  # add a "skill" to the robots skillset the control system will send a string with the ls_item and action and here we will look if we have a matching skill to execute
  # the item_modell defines the patterns which have to be used by the robot on multiple racks and or multiple samples in a rackpattern
  # inner pattern is always dependung on the object that has to be moved and the outer pattern is the pattern for the containers where the objects are stored in.
  # if racks have to be handled it is also an inner pattern cause the object to handle is the rack itself
  # create_item(id=0, ls_item="default", frame=p[0,0,0,0,0,0], actionlist=create_action_list([]), item_model=create_item_model(), lm_id=0, description="default")
  # create_item_model(inner=create_pattern(), outer=create_pattern(), description="default")
  # ITEM_MAP.append(create_item(id=1, ls_item="Home", frame=F1_uLM_Home, actionlist=[ActionManipulator.MOVE_TO], description="uLM Move To Home"))
  # ITEM_MAP.append(create_item(id=2, ls_item="InputStation", frame=F2_uLM_Input, actionlist=[ActionManipulator.PICK, ActionManipulator.PLACE], item_model=create_item_model(inner=Patterns.INPUT), description="uLM Pick and Place samples from Input"))
  # ITEM_MAP.append(create_item(id=3, ls_item="InputCapture", frame=F3_Cap_Input, actionlist=[ActionCamera.INSPECT, ActionManipulator.MOVE_TO], description="uLM Inspect samples from Input and Move To Capture Position"))
  # ITEM_MAP.append(create_item(id=4, ls_item="Bin", frame=F4_uLM_Bin, actionlist=[ActionManipulator.PLACE], description="uLM Place Cap to Bin"))
  # ITEM_MAP.append(create_item(id=5, ls_item="StationaryGripper", frame=F5_uLM_Gripper, actionlist=[ActionManipulator.PICK, ActionManipulator.PLACE, ActionManipulator.DECAP, ActionManipulator.MOVE_TO, ActionManipulator.GRASP, ActionManipulator.RELEASE], description=" uLM stationary gripper"))
  # ITEM_MAP.append(create_item(id=6, ls_item="CobasRack", frame=F6_uLM_Cobas_R, actionlist=[ActionManipulator.PICK, ActionManipulator.PLACE], item_model=create_item_model(outer=Patterns.COBAS_MAGAZINE), description="uLM Cobas Racks Pick and Place"))
  # ITEM_MAP.append(create_item(id=7, ls_item="CobasMagazine", frame=F7_uLM_Coba_Mag, actionlist=[ActionManipulator.PICK, ActionManipulator.PLACE], item_model=create_item_model(inner=Patterns.COBAS, outer=Patterns.COBAS_MAGAZINE), description="uLM Cobas Magazine Samples Pick and Place"))
  # ITEM_MAP.append(create_item(id=8, ls_item="DetectCobasRacks", frame=F8_Cap_Cobas_LM, actionlist=[ActionCamera.DETECT_OBJECTS, ActionManipulator.MOVE_TO], lm_id=2, description="uLM Cobas Rack Detection and Move To Capture"))
  # ITEM_MAP.append(create_item(id=9, ls_item="TaraMagazine", frame=F9_uLM_Tara, actionlist=[ActionManipulator.PICK, ActionManipulator.PLACE], item_model=create_item_model(inner=Patterns.TARA), description="uLM Centrifuge Tara Pick and Place"))
  # ITEM_MAP.append(create_item(id=10, ls_item="CentrifugeCapture", frame=F10_Cap_CF, actionlist=[ActionManipulator.MOVE_TO, ActionCamera.DETECT], lm_id=1, description="Centrifuge Device Move to Capture Pos and Detect Landmarks"))
  # ITEM_MAP.append(create_item(id=11, ls_item="Centrifuge", frame=F11_CF_PiPl, actionlist=[ActionManipulator.PICK, ActionManipulator.PLACE], description="Centrifuge Device Rack Pick and Place"))
  # ITEM_MAP.append(create_item(id=12, ls_item="CentrifugeMagazine", frame=F12_uLM_CF_Mag, actionlist=[ActionManipulator.PICK, ActionManipulator.PLACE], item_model=create_item_model(inner=Patterns.CENTRIFUGE, outer=Patterns.CENTRIFUGE_MAGAZINE), description=" uLM Centrifuge Magazin Pick and Place"))
  # ITEM_MAP.append(create_item(id=13, ls_item="CentrifugeRack", frame=F13_uLM_CF_R, actionlist=[ActionManipulator.PICK, ActionManipulator.PLACE], item_model=create_item_model(outer=Patterns.CENTRIFUGE_MAGAZINE), description="uLM Centrifuge Magazin Pick and Place Racks"))
  # ITEM_MAP.append(create_item(id=14, ls_item="DailyArchive", frame=F14_uLM_Archive, actionlist=[ActionManipulator.PICK, ActionManipulator.PLACE], item_model=create_item_model(inner=Patterns.ARCHIVE), description="uLM Pick and Place samples from Archive Rack"))
  # ITEM_MAP.append(create_item(id=15, ls_item="NokRack", frame=F15_uLM_Nok, actionlist=[ActionManipulator.PICK, ActionManipulator.PLACE], item_model=create_item_model(inner=Patterns.NOK), description="uLM Pick and Place samples from Nok Rack"))
  # ITEM_MAP.append(create_item(id=16, ls_item="CobasInput", frame=F16_Cobas_Input, actionlist=[ActionManipulator.PLACE], description="uLM Place Cobasrack in Cobas Device"))
  # ITEM_MAP.append(create_item(id=17, ls_item="CobasInputCapture", frame=F17_Cobas_Cap, actionlist=[ActionCamera.DETECT, ActionManipulator.MOVE_TO], lm_id=3, description="uLM Place Cobasrack in Cobas Device"))
  # ITEM_MAP.append(create_item(id=18, ls_item="XN550Input", frame=F18_XN550_Input, actionlist=[ActionManipulator.PICK, ActionManipulator.PLACE], item_model=create_item_model(inner=Patterns.SYSMEX_XN550, outer=Patterns.DRAWER_XN550), lm_id=4, description="uLM Pick and Place Samples in or out of XN550 Racks"))
  # ITEM_MAP.append(create_item(id=19, ls_item="XN550Capture", frame=F19_XN550_Cap, actionlist=[ActionCamera.DETECT, ActionManipulator.MOVE_TO], lm_id=4, description="uLM Move To and Capture LM XN550"))
  # ITEM_MAP.append(create_item(id=20, ls_item="XN550Drawer", frame=F20_XN550_Draw, actionlist=[ActionManipulator.DRAWER_OPEN, ActionManipulator.DRAWER_CLOSE], item_model=create_item_model(inner=Patterns.DRAWER_XN550), lm_id=4, description="uLM Open and close Drawer XN550"))
  # ITEM_MAP.append(create_item(id=21, ls_item="XN550Button", frame=F21_XN550_Btn, actionlist=[ActionManipulator.PUSH], lm_id=4, description="uLM Push XN550 Button"))
  # ITEM_MAP.append(create_item(id=22, ls_item="AMR", frame=p[0,0,0,0,0,0], actionlist=[ActionAMR.READ, ActionAMR.LOAD_MISSION, ActionAMR.START_MISSION, ActionAMR.NAVIGATE, ActionAMR.ACKNOWLEDGE], description="all AMR actions"))



  # ITEM_MAP.append(create_item(id=31, ls_item="TestLM", frame=TestLM, actionlist=[ActionManipulator.PICK, ActionManipulator.PLACE], item_model=create_item_model(inner=Rack.SYSMEX_CS2500), lm_id=5, description="LM Test"))
  # Fills the Vision Config List with Projectrelated Data
  # workspaceid and skillid are highly robominds related so probably will not stay like this in the future
  # sample detection: dx and dy are used to calculate the positions in a rack and given by the offset which will be applied in order to assign the sample to a place in the rack
  # create_vision_config(workspace_id="", skill_id="", item_id=-1, capture_pos=p[0,0,0,0,0,0], dx=0, dy=0, target_origin=p[0,0,0,0,0,0], selector="default", description="default")
  # VISION_CONFIG_MAP.append(create_vision_config(workspace_id="96017791-f581-4e9e-93da-6951695fccc8", skill_id="8885cfe1-6784-4293-bd26-52ebdc67bf95", capture_pos=F10_Cap_CF, target_origin=p[0,0,0,0,0,0], item_id=11, description="LM Detect CF"))
  # VISION_CONFIG_MAP.append(create_vision_config(workspace_id="96017791-f581-4e9e-93da-6951695fccc8", skill_id="8885cfe1-6784-4293-bd26-52ebdc67bf95", capture_pos=F8_Cap_Cobas_LM, target_origin=p[0,0,0,0,0,0], item_id=8, description="LM Detect Cobas Racks"))
  # VISION_CONFIG_MAP.append(create_vision_config(workspace_id="8f0ad01c-dc36-4fdd-b295-0b6b4a38b89a", skill_id="afdc9e13-ea83-40d6-a805-bb041453d2e5", capture_pos=F3_Cap_Input, target_origin=F2_uLM_Input, item_id=3, description="Lab Solution Input Capture"))
  # VISION_CONFIG_MAP.append(create_vision_config(workspace_id="96017791-f581-4e9e-93da-6951695fccc8", skill_id="8885cfe1-6784-4293-bd26-52ebdc67bf95", capture_pos=F19_XN550_Cap, target_origin=F18_XN550_Input, item_id=18, description="Input XN550"))
  # VISION_CONFIG_MAP.append(create_vision_config(workspace_id="96017791-f581-4e9e-93da-6951695fccc8", skill_id="8885cfe1-6784-4293-bd26-52ebdc67bf95", capture_pos=F19_XN550_Cap, target_origin=POS_Z, item_id=19, description="LM Detect XN550F"))
  # VISION_CONFIG_MAP.append(create_vision_config(workspace_id="96017791-f581-4e9e-93da-6951695fccc8", skill_id="8885cfe1-6784-4293-bd26-52ebdc67bf95", capture_pos=F10_Cap_CF, target_origin=POS_Z, item_id=10, description="LM Detect CF"))
  # VISION_CONFIG_MAP.append(create_vision_config(workspace_id="96017791-f581-4e9e-93da-6951695fccc8", skill_id="8885cfe1-6784-4293-bd26-52ebdc67bf95", capture_pos=F19_XN550_Cap, target_origin=F20_XN550_Draw, item_id=20, description="Drawer XN550"))
  # VISION_CONFIG_MAP.append(create_vision_config(workspace_id="96017791-f581-4e9e-93da-6951695fccc8", skill_id="8885cfe1-6784-4293-bd26-52ebdc67bf95", capture_pos=F19_XN550_Cap, target_origin=F21_XN550_Btn, item_id=21, description="Button XN550"))
  # VISION_CONFIG_MAP.append(create_vision_config(workspace_id="96017791-f581-4e9e-93da-6951695fccc8", skill_id="8885cfe1-6784-4293-bd26-52ebdc67bf95", capture_pos=TestLMCap, target_origin=p[0,0,0,0,0,0], item_id=30, description="Button XN550"))
  # VISION_CONFIG_MAP.append(create_vision_config(workspace_id="96017791-f581-4e9e-93da-6951695fccc8", skill_id="8885cfe1-6784-4293-bd26-52ebdc67bf95", capture_pos=TestLMCap, target_origin=TestLM, item_id=31, description="Button XN550"))

  # VISION_CONFIG_MAP.append(create_vision_config(workspace_id="96017791-f581-4e9e-93da-6951695fccc8", skill_id="8885cfe1-6784-4293-bd26-52ebdc67bf95", target_origin=p[0,0,0,0,0,0], item_id=11, description="LM Detect CF"))
  # VISION_CONFIG_MAP.append(create_vision_config(workspace_id="96017791-f581-4e9e-93da-6951695fccc8", skill_id="8885cfe1-6784-4293-bd26-52ebdc67bf95", target_origin=p[0,0,0,0,0,0], item_id=8, description="LM Detect Cobas Racks"))
  # VISION_CONFIG_MAP.append(create_vision_config(workspace_id="8f0ad01c-dc36-4fdd-b295-0b6b4a38b89a", skill_id="afdc9e13-ea83-40d6-a805-bb041453d2e5", target_origin=F2_uLM_Input, item_id=3, description="Lab Solution Input Capture"))
  # VISION_CONFIG_MAP.append(create_vision_config(workspace_id="96017791-f581-4e9e-93da-6951695fccc8", skill_id="8885cfe1-6784-4293-bd26-52ebdc67bf95", target_origin=F18_XN550_Input, item_id=18, description="Input XN550"))
  # VISION_CONFIG_MAP.append(create_vision_config(workspace_id="96017791-f581-4e9e-93da-6951695fccc8", skill_id="8885cfe1-6784-4293-bd26-52ebdc67bf95", target_origin=POS_Z, item_id=19, description="LM Detect XN550F"))
  # VISION_CONFIG_MAP.append(create_vision_config(workspace_id="96017791-f581-4e9e-93da-6951695fccc8", skill_id="8885cfe1-6784-4293-bd26-52ebdc67bf95", target_origin=POS_Z, item_id=10, description="LM Detect CF"))
  # VISION_CONFIG_MAP.append(create_vision_config(workspace_id="96017791-f581-4e9e-93da-6951695fccc8", skill_id="8885cfe1-6784-4293-bd26-52ebdc67bf95", target_origin=F20_XN550_Draw, item_id=20, description="Drawer XN550"))
  # VISION_CONFIG_MAP.append(create_vision_config(workspace_id="96017791-f581-4e9e-93da-6951695fccc8", skill_id="8885cfe1-6784-4293-bd26-52ebdc67bf95", target_origin=F21_XN550_Btn, item_id=21, description="Button XN550"))
  # VISION_CONFIG_MAP.append(create_vision_config(workspace_id="96017791-f581-4e9e-93da-6951695fccc8", skill_id="8885cfe1-6784-4293-bd26-52ebdc67bf95", target_origin=p[0,0,0,0,0,0], item_id=30, description="Button XN550"))
  # VISION_CONFIG_MAP.append(create_vision_config(workspace_id="96017791-f581-4e9e-93da-6951695fccc8", skill_id="8885cfe1-6784-4293-bd26-52ebdc67bf95", target_origin=TestLM, item_id=31, description="Button XN550"))

  # local inputrack = find_pattern_by_name("INPUT")
  # INSPECT_CONFIG_MAP.append(create_inspect_config(item_id=3, dx=inputrack.pattern_width[0]/(inputrack.pattern_size[0]-1), dy=inputrack.pattern_width[1]/(inputrack.pattern_size[1]-1), rack_size=inputrack.pattern_size , description="Input Capture"))
  # # Fills the Landmark List with Projectrelated Data
  # # create_landmark(lm_id=0, marker_id=-1, marker_size=0.1, marker_type="aruco_7x7", capture_pos=p[0,0,0,0,0,0], init_frame=p[0,0,0,0,0,0], search_offset=[0,0,0], actual_frame=p[0,0,0,0,0,0], description="")
  # LANDMARK_MAP.append(create_landmark(lm_id=1, marker_id=3, marker_size=0.1, marker_type="aruco_7x7", capture_pos = F10_Cap_CF, init_frame=p[-0.617789, -0.065471, 0.07918, 0.020983, -0.012695, 1.512066], search_offset=[0.15, 0.15, 0.1], actual_frame=p[-0.617789, -0.065471, 0.07918, 0.020983, -0.012695, 1.512066], description="LM CF Lid"))
  # LANDMARK_MAP.append(create_landmark(lm_id=2, marker_id=-1, marker_size=0.0085, marker_type="aruco_4x4", capture_pos = F8_Cap_Cobas_LM, init_frame=p[0,0,0,0,0,0], search_offset=[0.15, 0.15, 0.1], actual_frame=POS_Z, description="LM Cobas Rack Detection"))
  # LANDMARK_MAP.append(create_landmark(lm_id=3, marker_id=0, marker_size=0.1, marker_type="aruco_7x7", capture_pos = F17_Cobas_Cap, init_frame=p[-0.667,-0.194,0.100,0,0,0], search_offset=[0.15, 0.15, 0.1], actual_frame=POS_Z, description="LM Cobas Cap"))
  # LANDMARK_MAP.append(create_landmark(lm_id=4, marker_id=4, marker_size=0.1, marker_type="aruco_7x7", capture_pos = F19_XN550_Cap, init_frame=p[0.124,-0.976,0.355,-0.008,0.025,3.131], search_offset=[0.15, 0.15, 0.1], actual_frame=p[0,0,0,0,0,0], description="LM XN550 Cap"))
  # LANDMARK_MAP.append(create_landmark(lm_id=5, marker_id=0, marker_size=0.1, marker_type="aruco_7x7", capture_pos = TestLMCap, init_frame=p[-0.49,-0.144,0.092,0,-0.008,0.001], search_offset=[0.15, 0.15, 0.1], actual_frame=POS_Z, description="LM Test"))
  # # Configuration of all movement related parameters
  # # create_movement(id=0, hh_approach=POS_Z, h_approach=POS_Z, approach=POS_Z, h_target=POS_Z, target=POS_Z, retract=POS_Z, h_retract=POS_Z, hh_retract=POS_Z, h_frame=POS_Z, frame=POS_Z, speed=1, acceleration=1, description="default")
  # MOVEMENT_MAP.append(create_movement(description="TestLMCap", frame=TestLMCap, actionlist=[ActionManipulator.MOVE_TO]))
  # MOVEMENT_MAP.append(create_movement(description="TestLM", frame=TestLM, actionlist=[ActionManipulator.PICK,ActionManipulator.PLACE],
  #         approach=p[0,0,0.1,0,0,0],
  #         retract=p[0,0,0.1,0,0,0]))
  # MOVEMENT_MAP.append(create_movement(description="Home - MOVE_TO", frame=F1_uLM_Home, actionlist=[ActionManipulator.MOVE_TO]))
  # MOVEMENT_MAP.append(create_movement(description="Input - PICK&PLACE", frame=F2_uLM_Input, actionlist=[ActionManipulator.PICK,ActionManipulator.PLACE],
  #         approach=p[0,0,0.1,0,0,0],
  #         retract=p[0,0,0.1,0,0,0]))
  # MOVEMENT_MAP.append(create_movement(description="Capture Input - MOVE_TO", frame=F3_Cap_Input, actionlist=[ActionManipulator.MOVE_TO]))
  # MOVEMENT_MAP.append(create_movement(description="BIN - PLACE", frame=F4_uLM_Bin, actionlist=[ActionManipulator.PLACE],
  #         approach=p[0,0,0.1,0,0,0],
  #         retract=p[0,0,0.1,0,0,0]))
  # MOVEMENT_MAP.append(create_movement(description="Gripper - Move To", frame=F5_uLM_Gripper, actionlist=[ActionManipulator.MOVE_TO],
  #         approach=p[0,0,0.1,0,0,0]))
  # MOVEMENT_MAP.append(create_movement(description="Gripper - Pick", frame=F5_uLM_Gripper, actionlist=[ActionManipulator.PICK],
  #         retract=p[0,0,0.1,0,0,0]))
  # MOVEMENT_MAP.append(create_movement(description="Gripper - Place", frame=F5_uLM_Gripper, actionlist=[ActionManipulator.PLACE],
  #         approach=p[0,0,0.1,0,0,0]))
  # MOVEMENT_MAP.append(create_movement(description="CobasRack Pick & Place", frame=F6_uLM_Cobas_R, actionlist=[ActionManipulator.PICK,ActionManipulator.PLACE],
  #         approach=p[0,0,0.1,0,0,0],
  #         target=p[0,0,0,0,0,d2r(90)],
  #         retract=p[0,0,0.1,0,0,0]))
  # MOVEMENT_MAP.append(create_movement(description="CobasMagazine Pick & Place", frame=F7_uLM_Coba_Mag, actionlist=[ActionManipulator.PICK,ActionManipulator.PLACE],
  #         approach=p[0,0,0.1,0,0,0],
  #         target=p[0,0,0,0,0,-d2r(90)],
  #         retract=p[0,0,0.1,0,0,0]))
  # MOVEMENT_MAP.append(create_movement(description="Capture Position Cobas Landmarks", frame=F8_Cap_Cobas_LM, actionlist=[ActionManipulator.MOVE_TO]))
  # MOVEMENT_MAP.append(create_movement(description="TaraMagazine - PICK & PLACE", frame=F9_uLM_Tara, actionlist=[ActionManipulator.PICK,ActionManipulator.PLACE],
  #         approach=p[0,0,0.13,0,0,0],
  #         target=p[0,0,0,0,0,-d2r(90)],
  #         retract=p[0,0,0.13,0,0,0]))
  # MOVEMENT_MAP.append(create_movement(description="Capture Position - Centrifuge LM", frame=F10_Cap_CF,actionlist=[ActionManipulator.MOVE_TO]))
  # MOVEMENT_MAP.append(create_movement(description="Pick and Place Racks - Centrifuge Lid", frame=F11_CF_PiPl, actionlist=[ActionManipulator.PICK,ActionManipulator.PLACE],
  #         approach=p[0,0,0.3,0,0,0],
  #         retract=p[0,0,0.3,0,0,0]))
  # MOVEMENT_MAP.append(create_movement(description="Pick and Place Samples - Centrifuge on uLM", frame=F12_uLM_CF_Mag, actionlist=[ActionManipulator.PICK,ActionManipulator.PLACE],
  #         approach=p[0,0,0.13,0,0,0],
  #         retract=p[0,0,0.13,0,0,0]
  #         ))
  # MOVEMENT_MAP.append(create_movement(description="Pick and Place Racks - Centrifuge on uLM", frame=F13_uLM_CF_R, actionlist=[ActionManipulator.PICK,ActionManipulator.PLACE],
  #         approach=p[0,0,0.15,0,0,0],
  #         retract=p[0,0,0.15,0,0,0]
  #         ))

  # MOVEMENT_MAP.append(create_movement(description="Pick and Place Samples XN550 Racks in Device", frame=F18_XN550_Input, actionlist=[ActionManipulator.PICK,ActionManipulator.PLACE],
  #         approach=p[0,0,0.1,0,0,0],
  #         target = p[0,0,0,0,0,d2r(90)],
  #         retract=p[0,0,0.1,0,0,0]
  #         ))
  # MOVEMENT_MAP.append(create_movement(description="Capture LM XN550", frame=F19_XN550_Cap, actionlist=[ActionManipulator.MOVE_TO]))
  # MOVEMENT_MAP.append(create_movement(description="Open XN550 Drawer ", frame=F20_XN550_Draw, actionlist=[ActionManipulator.DRAWER_OPEN],
  #         h_approach=p[0.07,0,0.1,0,0,0],
  #         approach=p[0,0,0.1,0,0,0],
  #         target = p[0,0,0,0,0,d2r(90)],
  #         retract=p[0.07,0,0,0,0,0],
  #         h_retract=p[0.07,0,0.1,0,0,0]
  #         ))
  # MOVEMENT_MAP.append(create_movement(description="Close XN550 Drawer ", frame=F20_XN550_Draw, actionlist=[ActionManipulator.DRAWER_CLOSE],
  #         h_approach=p[0.07,0,0.1,0,0,0],
  #         approach=p[0.07,0,0,0,0,0],
  #         target = p[0,0,0,0,0,d2r(90)],
  #         retract=p[0,0,0.1,0,0,0],
  #         h_retract=p[0.07,0,0.1,0,0,0]
  #         ))
  # MOVEMENT_MAP.append(create_movement(description="Push XN550 Button ", frame=F21_XN550_Btn, actionlist=[ActionManipulator.PUSH],
  #         approach=p[0,0,0.15,0,0,0],
  #         retract=p[0,0,0.15,0,0,0]
  #         ))
  # MOVEMENT_MAP.append(create_movement(description="Capture Position 2 Input", frame=F_Cap_Input2,actionlist=[ActionManipulator.MOVE_TO]))



  $ 19 "Script: SCRIPT Objects V0.1.script"
  #*****************************************************
  # customer          :   INTERNAL
  # project name      :
  #****************************************************
  # controller        :   UR
  # software          :   5.17.3
  #****************************************************
  # author            :   P. Koehnke
  # Copyright (c)     :   United Robotics Group
  #                       An der Riede 2
  #                       28816 Stuhr
  #                       Germany
  #****************************************************
  # description       :   object database
  # version:      	:   0.1
  # created           :   09.10.2024
  # updated           :
  #****************************************************
  # modifications     :
  #
  # date              :
  # name              :
  # reason            :
  #****************************************************

  def create_object_2(id=0, name="", type=0, dimension=struct(length=0, width=0, height=0, diameter=0), gripper_offset=p[0,0,0,0,0,0]):
      return struct(id=id, name=name, type=type, dimension=dimension, gripper_offset=gripper_offset)
  end

  OBJ = create_object_2()
  OBJs = make_list(0, create_object_2(), 50)

  OBJs.append(create_object_2(id=1, name="rack centrifuge", type=1, dimension=struct(length=0, width=0, height=0.106, diameter=0.020), gripper_offset=p[0,0,0.095,0,0,2.356]))
  OBJs.append(create_object_2(id=2, name="sample tube 1", type=2, dimension=struct(length=0, width=0, height=0.106, diameter=0.015), gripper_offset=p[0,0,0,0,0,0]))
  OBJs.append(create_object_2(id=3, name="rack sarstedt", type=3, dimension=struct(length=0, width=0, height=0.100, diameter=0.020), gripper_offset=p[0,0,0,0,0,0]))
  OBJs.append(create_object_2(id=4, name="Lab bottle", type=4, dimension=struct(length=0, width=0, height=0.100, diameter=0.030), gripper_offset=p[0,0,0.2,0,0,0]))
  OBJs.append(create_object_2(id=5, name="Vial", type=5, dimension=struct(length=0, width=0, height=0.100, diameter=0.0275), gripper_offset=p[0,0,0,0,0,0]))
  OBJs.append(create_object_2(id=6, name="Container", type=6, dimension=struct(length=0.09, width=0.09, height=0.185, diameter=0.080), gripper_offset=p[0,0,0,0,0,0]))
  OBJs.append(create_object_2(id=7, name="Target_container", type=7, dimension=struct(length=0.06, width=0.06, height=0.134, diameter=0.05), gripper_offset=p[0,0,0,0,0,0]))
  OBJs.append(create_object_2(id=8, name="Spatula", type=8, dimension=struct(length=0.03, width=0.03, height=0.23, diameter=0.05), gripper_offset=p[0,0,0,0,0,0]))
  OBJs.append(create_object_2(id=9, name="rack pipet", type=9, dimension=struct(length=0.03, width=0.03, height=0.23, diameter=0.05), gripper_offset=p[0,0,0,0,0,0]))

  def create_jig_2(id=0, name="", type=0, capacity=0, jig_offset=p[0,0,0,0,0,0]):
      # iformation about used jigs
      return struct(id=id, name=name, type=type, capacity=capacity, jig_offset=jig_offset)
  end

  JIG2 = create_jig_2()
  JIGs = make_list(0, create_jig_2(), 20)

  JIGs.append(create_jig_2(id=1, name="3FG", type=1, capacity=1, jig_offset=p[0,0,0,0,0,0]))
  JIGs.append(create_jig_2(id=2, name="jig input", type=2, capacity=1, jig_offset=p[0,0,0,0,0,-3.927]))
  JIGs.append(create_jig_2(id=3, name="jig output", type=3, capacity=1, jig_offset=p[0,0,0,0,0,0.78]))
  JIGs.append(create_jig_2(id=6, name="jig bin", type=6, capacity=1, jig_offset=p[0,0,0,0,0,0]))
  JIGs.append(create_jig_2(id=7, name="jig sarstedt racks", type=7, capacity=1, jig_offset=p[0,0,-0.02,0,0,0]))
  JIGs.append(create_jig_2(id=8, name="NoK Bin", type=8, capacity=1, jig_offset=p[0,0,0,0,0,0]))
  JIGs.append(create_jig_2(id=9, name="Pick bott jig", type=9, capacity=1, jig_offset=p[0,0,0,0,0,0]))
  JIGs.append(create_jig_2(id=10, name="Place bott jig", type=10, capacity=1, jig_offset=p[0,0,0,0,0,0]))
  JIGs.append(create_jig_2(id=11, name="bottle shake jig", type=11, capacity=1, jig_offset=p[0,0,0,0,0,0]))
  JIGs.append(create_jig_2(id=12, name="Pick Vial jig", type=12, capacity=1, jig_offset=p[0,0,0,0,0,0]))
  JIGs.append(create_jig_2(id=13, name="Place Vial jig", type=13, capacity=1, jig_offset=p[0,0,0,0,0,0]))
  JIGs.append(create_jig_2(id=14, name="Liquid transfer jig", type=14, capacity=1, jig_offset=p[0,0,0,0,0,0]))
  JIGs.append(create_jig_2(id=15, name="Pick station jig", type=15, capacity=1, jig_offset=p[0,0,0,0,0,0]))
  JIGs.append(create_jig_2(id=16, name="Place station jig", type=16, capacity=1, jig_offset=p[0,0,0,0,0,0]))
  JIGs.append(create_jig_2(id=17, name="Weigh station jig", type=17, capacity=1, jig_offset=p[0,0,0,0,0,0]))
  JIGs.append(create_jig_2(id=18, name="Pick station 1", type=18, capacity=1, jig_offset=p[0,0,0,0,0,0]))
  JIGs.append(create_jig_2(id=19, name="Pick station 2", type=19, capacity=1, jig_offset=p[0,0,0,0,0,0]))
  JIGs.append(create_jig_2(id=20, name="Pick station 3", type=20, capacity=1, jig_offset=p[0,0,0,0,0,0]))
  JIGs.append(create_jig_2(id=21, name="Tilt station jig", type=21, capacity=1, jig_offset=p[0,0,0,0,0,0]))
  $ 20 "Script: Tilting.script"
  global g_has_ref = False
  global g_pivot_pose = p[0, 0, 0, 0, 0, 0]
  global g_rel0 = p[0, 0, 0, 0, 0, 0]
  global g_current_angle = 0.0

  hinge_offset = p[0, 0, -0.20, 0, 0, 0]
  global g_rq_ready = False
  global RQ_FORCE = 30
  global RQ_SPEED = 100
  global RQ_GRIP_TIMEOUT = 2.0

  def tilt_init_reference():
  	p_center = get_actual_tcp_pose()
  	g_pivot_pose = pose_trans(p_center, hinge_offset)
  	g_rel0 = pose_trans(pose_inv(g_pivot_pose), p_center)
  	g_current_angle = 0.0
  	g_has_ref = True
  end

  def rq_ensure_ready():
  	if (not g_rq_ready):
  		rq_activate_and_wait()
  		rq_set_force(RQ_FORCE)
  		rq_set_speed(RQ_SPEED)
  		g_rq_ready = True
  	end
  end



  #def rq_open_and_wait():
  	#rq_open()
  	#sleep(0.25)
  #end

  def tilt_to(target_deg):
  	if ( not g_has_ref):
  		tilt_init_reference()
  	end

  	rq_ensure_ready()
  	rq_close_and_wait()

  	angle_mid = (g_current_angle + target_deg)/2.0
  	rad_mid = (angle_mid)*3.1416/180
  	rad_end = target_deg*3.1416/180

  	tilt_mid = p[0,0,0, -rad_mid, 0, 0]
  	tilt_end = p[0,0,0, -rad_end, 0, 0]

  	pose_rel_mid = pose_trans(tilt_mid, g_rel0)
  	pose_rel_end = pose_trans(tilt_end, g_rel0)

  	via_pose = pose_trans(g_pivot_pose, pose_rel_mid)
  	end_pose = pose_trans(g_pivot_pose, pose_rel_end)

  	movec(via_pose, end_pose, a=0.05, v=0.01, r=0.001)

  	rq_open_and_wait()

  	g_current_angle = target_deg
  end


  def tilt_by(delta_deg):
  	tilt_to(g_current_angle + delta_deg)
  end

  def tilt_reset():
  	g_has_ref = False
  end

  $ 21 "Script: recipe_updated.script"
  # ============================================
  # Recipe Dosing URScript (3 powders, sorted A/B/C)
  # - keeps final mixture ratio after 1st overshoot
  # - syncs with Python dashboard via TCP
  # ============================================

  # --------- HANDOFF GLOBALS (used by other skills) ---------
  global Pow_name = ""
  global target_weight = 0.0
  global last_dose_error = 0.0

  # --------- RECIPE STATE ---------
  global powder_names = ["", "", ""]
  global powder_ratios = [0.0, 0.0, 0.0]      # fractions 0..1
  global powder_targets = [0.0, 0.0, 0.0]     # target weights for each powder
  global powder_actuals = [0.0, 0.0, 0.0]     # measured after dosing
  global powder_order  = [0, 1, 2]            # indices, sorted by ascending ratio

  global total_weight = 0.0                   # initial / adjusted total
  global current_powder_index = 0             # index into powder_order
  global ratio_adjusted = False               # did we already adjust after powder 1
  global dose_start_weight = 0.0              # weight at dosing start for each powder

  # --------- FINAL RESULTS (for dashboard) ---------
  # WA/WB/WC = final weights of powders A/B/C after dosing (sorted by ratio)
  global WA = 0.0
  global WB = 0.0
  global WC = 0.0

  # finalPercA/B/C = final percentages of WA/WB/WC wrt adjusted total
  global finalPercA = 0.0
  global finalPercB = 0.0
  global finalPercC = 0.0

  # counter to know which powder we just finished (1 → A, 2 → B, 3 → C)
  global dose_counter = 0


  # =====================================================
  # SORTING HELPERS (BY ASCENDING RATIO)
  # =====================================================

  def swap_order(i, j):
    local temp = powder_order[i]
    powder_order[i] = powder_order[j]
    powder_order[j] = temp
  end

  def sort_powders_by_ratio():
    # bubble-sort style, only 3 elements
    global powder_order = [0, 1, 2]

    if (powder_ratios[powder_order[1]] < powder_ratios[powder_order[0]]):
      swap_order(0, 1)
    end

    if (powder_ratios[powder_order[2]] < powder_ratios[powder_order[1]]):
      swap_order(1, 2)
    end

    if (powder_ratios[powder_order[1]] < powder_ratios[powder_order[0]]):
      swap_order(0, 1)
    end
  end


  # =====================================================
  # TCP SENDING HELPERS (Python dashboard @ 192.168.12.103:3002)
  # =====================================================

  # Send powder labels in sorted A/B/C order
  # A = least %, B = middle %, C = highest %
  def send_powder_labels():
    local A = powder_names[powder_order[0]]
    local B = powder_names[powder_order[1]]
    local C = powder_names[powder_order[2]]

    socket_open("192.168.12.103", 3002)
    local cmd = "SET_LABELS:" + A + ";" + B + ";" + C
    textmsg("Sending labels: ", cmd)
    socket_send_string(cmd)
    sleep(0.2)
    socket_close()
  end

  # Send initial recipe (TOTAL;PA;PB;PC) in sorted order
  # powder_ratios are fractions (0..1), we convert to %
  def send_init_recipe(total_w):
    local rA = powder_ratios[powder_order[0]] * 100
    local rB = powder_ratios[powder_order[1]] * 100
    local rC = powder_ratios[powder_order[2]] * 100

    socket_open("192.168.12.103", 3002)
    local cmd = "SET_INIT:" +
                to_str(total_w) + ";" +
                to_str(rA) + ";" +
                to_str(rB) + ";" +
                to_str(rC)
    textmsg("Sending INIT: ", cmd)
    socket_send_string(cmd)
    sleep(0.2)
    socket_close()
  end

  # Send final recipe:
  # SET_FINAL:ADJ_TOTAL;PA;PB;PC;WA;WB;WC
  # where PA/B/C = finalPercA/B/C, WA/B/C = final weights, adj_total = total_weight
  def send_final_recipe(adj_total):
    socket_open("192.168.12.103", 3002)

    local cmd = "SET_FINAL:" +
                to_str(adj_total) + ";" +
                to_str(finalPercA) + ";" +
                to_str(finalPercB) + ";" +
                to_str(finalPercC) + ";" +
                to_str(WA) + ";" +
                to_str(WB) + ";" +
                to_str(WC)
    textmsg("Sending FINAL: ", cmd)
    socket_send_string(cmd)
    sleep(0.2)
    socket_close()
  end


  # =====================================================
  # FINAL WEIGHT & PERCENTAGE LOGIC
  # =====================================================

  # Call this ONCE after each powder dosing is finished
  # final_weight = w_dosed_total of the just-finished powder
  def record_final_weight_for_current_powder(final_weight):
    dose_counter = dose_counter + 1

    if dose_counter == 1:
      WA = final_weight
      textmsg("Assigned WA (Powder A): ", WA)
    elif dose_counter == 2:
      WB = final_weight
      textmsg("Assigned WB (Powder B): ", WB)
    elif dose_counter == 3:
      WC = final_weight
      textmsg("Assigned WC (Powder C): ", WC)
    else:
      textmsg("WARNING: dose_counter > 3, ignoring extra weight")
    end
  end

  # Compute final percentages from WA/WB/WC and adjusted total
  def compute_final_percentages(adj_total):
    if adj_total <= 0:
      textmsg("ERROR: adj_total <= 0, cannot compute final %")
    else:
      finalPercA = WA / adj_total * 100
      finalPercB = WB / adj_total * 100
      finalPercC = WC / adj_total * 100
      textmsg("Final % A/B/C: ", finalPercA, finalPercB, finalPercC)
    end
  end


  # =====================================================
  # RECIPE INITIALIZATION
  # =====================================================

  # powA/B/C  : strings (e.g. "MCC", "CCS", "MAGNESIUM_STEARATE")
  # total     : initial total weight (g)
  # ratioA/B/C: fractions (0..1), e.g. 0.3, 0.2, 0.5
  def recipe_init(powA, powB, powC, total, ratioA, ratioB, ratioC):
    global powder_names  = [powA, powB, powC]
    global powder_ratios = [ratioA, ratioB, ratioC]
    global total_weight  = total

    global powder_targets = [total*ratioA, total*ratioB, total*ratioC]
    global powder_actuals = [0.0, 0.0, 0.0]

    global current_powder_index = 0
    global ratio_adjusted = False
    global dose_start_weight = 0.0

    dose_counter = 0
    WA = 0.0
    WB = 0.0
    WC = 0.0

    sort_powders_by_ratio()

    # NOTE: you call these from your main flow when you want:
    send_powder_labels()
    send_init_recipe(total)
  end


  # =====================================================
  # POSITION + CAMERA HELPERS (YOUR EXISTING LOGIC)
  # =====================================================

  def get_position_for_powder(Pow_name):
    if pos1_powder == Pow_name:
      return "Position1"
    elif pos2_powder == Pow_name:
      return "Position2"
    elif pos3_powder == Pow_name:
      return "Position3"
    else:
      return -1
    end
  end

  def extract_powder_name(raw_str):
    local idx_open  = str_find(raw_str, "(")
    local idx_close = str_find(raw_str, ")")

    if (idx_open < 0) or (idx_close < 0):
      return raw_str
    end

    local inside = ""
    local i = idx_open + 1
    while i < idx_close:
      inside = str_cat(inside, str_at(raw_str, i))
      i = i + 1
    end

    local idx_comma = str_find(inside, ",")
    if idx_comma < 0:
      return inside
    end

    local powder = ""
    local j = idx_comma + 1
    while j < str_len(inside):
      powder = str_cat(powder, str_at(inside, j))
      j = j + 1
    end

    return powder
  end

  def get_response_from_camera(target):
    movel(target, a=0.1, v=0.12, r=0)
    visor_trigger("1", "3.0", "arm")
    global response = visor_getResponse(1)
  end


  # =====================================================
  # RECIPE STEP SELECTION
  # =====================================================

  # Call recipe_next() before each dosing run.
  # Returns True if a powder exists, False if done.
  def recipe_next():
    if (current_powder_index >= 3):
      return False
    end

    local i = powder_order[current_powder_index]
    global Pow_name = powder_names[i]
    global target_weight = powder_targets[i]

    global powder_position = get_position_for_powder(Pow_name)

    if (Pow_name == "CCS"):
      W_now = 200.0
    elif (Pow_name == "MCC"):
      W_now = 131.0
    else:
      W_now = 100.0
    end

    return True
  end


  # =====================================================
  # DOSING START / END
  # =====================================================

  # Call at the beginning of each powder dosing run
  def dosing_start():
    global dose_start_weight = get_weight()
    global switch_spat_M = True
    global switch_spat_S = True
    global switch_spat_F_S = True
  end

  # Call after dosing is finished for current powder
  def dosing_end():
    local idx = powder_order[current_powder_index]
    local weight_after = get_weight()
    local actual_weight = weight_after - dose_start_weight

    # store actual weight
    local tmp = powder_actuals
    tmp[idx] = actual_weight
    global powder_actuals = tmp

    # save error
    global last_dose_error = actual_weight - powder_targets[idx]

    # store WA/WB/WC in dosing (sorted) order
    record_final_weight_for_current_powder(actual_weight)

    # one-time correction after first powder (ratio preserving)
    if ((current_powder_index == 0) and (not ratio_adjusted)):
      local j = powder_order[1]
      local k = powder_order[2]

      local ratio_first = powder_ratios[idx]
      if (ratio_first > 0.0):
        # new_total = actual / ratio_first
        local new_total = actual_weight / ratio_first
        if (new_total < 0.0):
          new_total = 0.0
        end

        local ttmp = powder_targets
        ttmp[idx] = actual_weight
        ttmp[j]   = new_total * powder_ratios[j]
        ttmp[k]   = new_total * powder_ratios[k]
        global powder_targets = ttmp

        global adj_total = new_total
      end

      global ratio_adjusted = True
    end

    global current_powder_index = current_powder_index + 1
  end

  $ 22 "Script: scooping.script"
  def scooping_init():
  	#global W_FULL = 300.010
  	global H_INNER = 0.15
  	global TCP_to_tip = 0.020
  	global depth_saftey = 0.005
  	global container_height = 0.120
  	global reach_margin = 0.03

  	global angle_min = 18.0
  	global angle_max = 68.0
  	global gain_per_percent = 0.5

  	global level_bias_below_center = 0.020

  	global level = 0.0
  	global tilt_angle_sent = 0.0
  	global w_dosed_total = 0.0
  	global last_scale = 0.0
  	global g_z0_hi = 0.01
  	global g_z100_hi = 0.10
  	global g_z_min = 0.018
  	global g_z_max = 0.150

  	#global g_exp = 0.80
  	#global g_k = 0.03
  	#global g_alpha = 0.7
  	global g_corr_max = 0.010

  	global g_prev_cum_w = -1.0
  	global g_depth_corr = 0.0
  	global spatula_len = 0.17
  	global target_g = 0.0
  	global scoop_ct = 0
  	global error_sum = 0.0
  	global error_sq_sum = 0.0
  	global scoop_g = 0.0
  	global w_dosed_total = 0.0

  	if (Pow_name=="NaCl"):
  		global W_FULL = 625.00
  		global g_exp = 0.80
  		global g_k = 0.03
  		global g_alpha = 0.7
  	elif (Pow_name == "Mannitol"):
  		global W_FULL = 300.00
  		global g_exp = 0.82
  		global g_k = 0.025
  		global g_alpha = 0.6
  	elif (Pow_name == "MCC"):
  		global W_FULL = 280.0
  		global g_exp = 0.82
  		global g_k = 0.035
  		global g_alpha = 0.7
  	elif (Pow_name == "CCS"):
  		global W_FULL = 250.0
  		global g_exp = 0.82
  		global g_k = 0.035
  		global g_alpha = 0.7
  	elif (Pow_name == "Magnesium_stearate"):
  		global W_FULL = 200.0
  		global g_exp = 0.84
  		global g_k = 0.025
  		global g_alpha = 0.6
  	elif (Pow_name == "lactose_fine"):
  		global W_FULL = 330.0
  		global g_exp = 0.84
  		global g_k = 0.025
  		global g_alpha = 0.55
  	else:
  		popup("Unkwon powder type. Using default NaCl settings.", title="Calibration Warning")
  		global W_FULL = 300.0
  		global g_k = 0.03
  		global g_alpha = 0.7
  	end


  end

  def clamp(x, lo, hi):
  	if(x<lo):
  		return lo
  	elif (x>hi):
  		return hi
  	else:
  		return x
  	end
  end

  def compute_level_percent(W_now, weight_value):
  	local delta = weight_value - last_scale
  	if (delta<0.0):
  		delta = 0.0
  	end
  	global w_dosed_total = w_dosed_total + delta
  	last_scale = weight_value

  	local W_eff = W_now-w_dosed_total
  	if (W_eff<W_EMPTY):
  		W_eff = W_EMPTY
  	end

  	level = 100.0* (W_eff -W_EMPTY)/ (W_FULL-W_EMPTY)
  	level = clamp(level,0.0,100.0)

  	return level
  end

  def compute_tilt_deg(level_percent):
  	angle = angle_min + gain_per_percent*(100.0-level_percent)
  	return clamp(angle, angle_min, angle_max)
  end


  def tilt(level_percentage):
  	new_angle = compute_tilt_deg(level_percentage)
  	global angle_rel = new_angle - tilt_angle_sent

  	if my_abs(angle_rel)>2.0:
  		tilt_send(new_angle)
  		global angle_deg = new_angle
  		global tilt_angle_sent = new_angle
  		global p_center = updated_center_pose(p_center_vertical, angle_deg)
  	end

  	if (level<85.0):
  		tilt_send(angle_deg)
  	end
  end

  def compute_scoop_depth(level, cum_w, target_g):
  	if (level >=10.0):
  		ratio = level/100.0
  		corrected = pow(ratio, g_exp)
  		base_z = g_z0_hi + (g_z100_hi - g_z0_hi)*corrected

  	elif (level<10.00 and level>=1.00):
  		z0 = 0.023
  		z100 = 0.140
  		ratio2 = level/100.0
  		base_z = z0 +(z100-z0)*ratio2
  	else:
  		base_z = 0.016
  	end

  	if (g_prev_cum_w<0):
  		g_prev_cum_w = cum_w

  	else:
  		global scoop_g = cum_w-g_prev_cum_w
  		g_prev_cum_w = cum_w

  		e = target_g -scoop_g

  		corr_proposed = g_k*e
  		g_depth_corr = (1.0 -g_alpha)*g_depth_corr + g_alpha*corr_proposed
  		g_depth_corr = clamp(g_depth_corr, -g_corr_max, g_corr_max)
  	end

  	z_tip = base_z - g_depth_corr
  	z_tip = clamp(z_tip, g_z_min, g_z_max)


  	return z_tip
  end

  def my_abs(val):
  	if (val<0):
  		return -val
  	else:
  		return val
  	end
  end


  def select_spatula(Pow_name, level, diff):
  	if (Pow_name == "lactose_fine" or Pow_name== "Magnesium_stearate"):
  		if (level >10.0 and diff>0.6):
  			return "spatula_flat_M"
  		else:
  			return "spatula_flat_S"
  		end

  	elif (Pow_name == "NaCl" and level >10.0 and diff>6.5):
  		return "spatula_L"
  	elif(Pow_name == "NaCl" and level> 10.0 and diff<=6.5):
  		return "spatula_M"
  	elif (Pow_name == "MCC" and level >10.0 and diff>2.0):
  		return "spatula_L"
  	elif(Pow_name == "MCC" and level> 10.0 and diff<=2.0):
  		return "spatula_M"
  	elif ((Pow_name == "Mannitol" or Pow_name == "CCS") and level >10.0 and diff>3.2):
  		return "spatula_L"
  	elif ((Pow_name == "Mannitol" or Pow_name == "CCS") and level >10.0 and diff<=3.2):
  		return "spatula_M"
  	elif( level>1.0 and level <= 10.0):
  		return "spatula_M"
  	else:
  		return "spatula_S"
  	end
  end

  global target_g_table = [
  	"NaCl", "spatula_L", "6.8",
  	"NaCl", "spatula_M", "1.75",
  	"NaCl", "spatula_S", "0.135",

  	"Mannitol", "spatula_L", "3.1",
  	"Mannitol", "spatula_M", "0.9",
  	"Mannitol", "spatula_S", "0.075",

  	"CCS", "spatula_L", "2.5",
  	"CCS", "spatula_M", "0.9",
  	"CCS", "spatula_S", "0.075",

  	"MCC", "spatula_L", "1.8",
  	"MCC", "spatula_M", "0.5",
  	"MCC", "spatula_S", "0.05",

  	"Magnesium_stearate", "spatula_flat_M", "0.5",
  	"Magnesium_stearate", "spatula_flat_S", "0.25",

  	"lactose_fine", "spatula_flat_M", "1.0",
  	"lactose_fine", "spatula_flat_S", "0.7"]

  def get_target_g(Pow_name, spat_name):
  	local i = 0
  	local n = length(target_g_table)
  	while (i < n):
  		if (target_g_table[i] == Pow_name and target_g_table[i+1] == spat_name):
  			return to_num(target_g_table[i+2])
  		end
  		i = i+3
  	end
  	popup("No target_g match for: ", Pow_name, ", ", spatula)

  end
  def auto_tilt_and_scoop(W_now, target_weight, weight_value):
  	level = compute_level_percent(W_now, weight_value)

  	global spatula = select_spatula(Pow_name, level, diff)
  	global target_g = get_target_g(Pow_name, spatula)

  	global scoop_depth = compute_scoop_depth(level, weight_value, target_g)

  	tilt(level)
  	#p_center = get_actual_tcp_pose()

  	if (scoop_ct < 5 and g_prev_cum_w>0.0):
  		#local scoop_g = scoop_g
  		local error = target_g - scoop_g
  		error_sum = error_sum + error
  		error_sq_sum = error_sq_sum + error*error
  		scoop_ct = scoop_ct+1

  		if (scoop_ct==5):
  			local avg_error = error_sum/5.0
  			#local std_dev = sqrt(error_sq_sum/5.0) - (avg_error*avg_error))

  			if (my_abs(avg_error)>1.0):
  				g_k = 0.055
  				g_alpha = 0.85
  			elif (my_abs(avg_error)>0.6):
  				g_k= 0.045
  				g_alpha =0.75
  			elif (my_abs(avg_error)> 0.3):
  				g_k = 0.035
  				g_alpha = 0.65
  			elif (my_abs(avg_error)>0.1):
  				g_k = 0.025
  				g_alpha = 0.55
  			else:
  				g_k = 0.015
  				g_alpha = 0.45
  			end
  		end
  	end

  	scoop_powder(p_center)
  end


  def after_scoop():
  	tilt_send(angle_deg)
  	sleep(0.5)
  	movel(lifted_pose, a=0.05, v=0.2)
  	movel(tilted_pose_in_base, a=0.05, v=0.2)
  	set_analog_out(0,0.4)
  	movel(pose_trans(tilted_pose_in_base, p[-0.01,0,0,0,0,2.0]), a=0.05, v=0.2)
  	set_analog_out(0,0.0)
  	movel(lifted_pose, a=0.05, v=0.2)
  	tilt_to_home()
  end
  $ 23 "Script: dosing.script"
  def vibration_2():
  	set_analog_out(0,0.4)
  	sleep(0.8)
  	set_analog_out(0,0.0)
  	sleep(0.2)
  end

  def vibration_3():
  	set_analog_out(0,0.4)
  	sleep(0.5)
  	set_analog_out(0,0.0)
  	sleep(0.3)
  end

  def vibration_4():
  	set_analog_out(0,0.4)
  	sleep(0.6)
  	set_analog_out(0, 0.0)
  	sleep(0.5)
  end

  def vibration_1():
  	set_analog_out(0,0.4)
  	sleep(1)
  	set_analog_out(0,0.0)
  	sleep(0)
  end

  def move_tilt_in_steps(Pow_center, final_pose, steps):
  	i = 0
  	while i <= steps:
  		ratio = i / steps
  		pose_step = p[Pow_center[0] + ratio * (final_pose[0] - Pow_center[0]), Pow_center[1] + ratio * (final_pose[1] -Pow_center[1]),Pow_center[2] + ratio * (final_pose[2] - Pow_center[2]), Pow_center[3] + ratio * (final_pose[3] - Pow_center[3]), Pow_center[4] + ratio * (final_pose[4] - Pow_center[4]), Pow_center[5] + ratio * (final_pose[5] - Pow_center[5])]
  		movej(pose_step, a=1.2, v=0.15)
  		sleep(0.1)
  		i = i+1
  	end
  end

  def tilt_container(angle):
  	p_center = get_actual_tcp_pose()
  	hinge_offset = p[0,0,-0.23,0,0,0]
  	pivot_pose = pose_trans(p_center, hinge_offset)
  	pose_rel = pose_trans(pose_inv(pivot_pose), p_center)
  	angle_mid = (angle/2.0)*3.1416/180
  	angle_end = angle*3.1416/180
  	tilt_mid = p[0,0,0, -angle_mid, 0, 0]
  	tilt_end = p[0,0,0, -angle_end, 0, 0]
  	pose_rel_mid = pose_trans(tilt_mid, pose_rel)
  	pose_rel_end = pose_trans(tilt_end, pose_rel)
  	via_pose = pose_trans(pivot_pose, pose_rel_mid)
  	end_pose = pose_trans(pivot_pose, pose_rel_end)
  	movec(via_pose, end_pose, a=0.05, v=0.01, r=0.001)
  	p_center = get_actual_tcp_pose()
  end

  def deg2rad(d):
  	return d*3.141592/180
  end

  def map_tilt_to_ry_deg(container_deg):
  	#ry_deg = -0.875*container_deg +87.0
  	#return clamp(ry_deg, 5.0, 80.0)
  	if (Pow_name == "NaCl" or Pow_name == "Mannitol" or Pow_name == "CCS" or Pow_name == "MCC"):
  		if ( level>=10.0):
  			ry_min = 10.0
  			ry_max = 75.0
  		elif (level<10.00 and level >1.00):
  			ry_min = 16.0
  			ry_max = 65.0
  		else:
  			ry_min=17.0
  			ry_max=75.0
  		end
  	else:
  		if ( level>=10.0):
  			ry_min = 0.0
  			ry_max = 65.0
  		elif (level<10.00 and level >1.00):
  			ry_min = 10.0
  			ry_max = 45.0
  		else:
  			ry_min=0.0
  			ry_max=50.0
  		end

  	end
  	local span_count = angle_max -angle_min
  	local span_ry = ry_max - ry_min

  	local t = (container_deg -angle_min)/span_count
  	local ry_deg = ry_max - t*span_ry

  	return clamp(ry_deg, ry_min, ry_max)

  end

  def caluclate_corrections(level):
  	z_high = 0.01
  	z_low = -0.08
  	y_high = -0.01
  	y_low = -0.015

  	scale = (level - 10.0) / (100.0-10.0)

  	global correction_z = z_low + scale*(z_high - z_low)
  	global correction_y = y_low + scale*(y_high -y_low)

  end

  def scoop_powder(p_center):
  	#lift_offset = p[0, 0, 0.05, 0, 0, 0]
  	vibration_voltage = 0.4
  	vibration_time = 3.0
  	diameter = 0.07
  	global scoop_radius_default = 0.0
  	#p_center = center_pose_t


  	if (level >=70.00):
  		approach_offset = p[0.008,0,0.22,0,0,0]
  		lift_offset = p[0, 0, 0.05, 0, 0, 0]
  		caluclate_corrections(level)
  	elif (level >=10.00 and level <70):
  		approach_offset = p[0.008,0,0.22,0,0,0]
  		lift_offset = p[0, 0, 0.15, 0, 0, 0]
  		caluclate_corrections(level)
  	elif (level<10.00 and level >= 1.00):
  		approach_offset = p[0.01,0,0.22,0,0,0]
  		correction_z = -0.08
  		correction_y = -0.01
  		lift_offset = p[0, 0, 0.14, 0, 0, 0]
  	else:
  		approach_offset = p[0.008,0,0.22,0,0,0]
  		correction_z = -0.08
  		correction_y = -0.01
  		lift_offset = p[0, 0, 0.14, 0, 0, 0]
   	end

  	if (spatula == "spatula_L"):
  		global spatula_depth = 0.015
  	elif (spatula == "spatula_M"):
  		global spatula_depth = 0.01
  	elif (spatula == "spatula_S"):
  		global spatula_depth = 0.008
  	elif (spatula == "spatula_flat_M"):
  		global spatula_depth = 0.001
  	elif (spatula == "spatula_flat_S"):
  		global spatula_depth = 0.005
  	end

  	scoop_radius_default = diameter/2 - spatula_depth
  	scoop_entry_pose = pose_trans(p_center, approach_offset)
  	movel(scoop_entry_pose, a=0.1, v=0.25)

  	scoop_start_rel = p[scoop_radius_default, 0, scoop_depth, 0, 0, 0]

  	rot_mid = p[0, 0, 0, 0, 0, 0.785]
  	rot_end = p[0, 0, 0, 0, 0, 1.5708]

  	scoop_via_rel = pose_trans(rot_mid, scoop_start_rel)
  	scoop_end_rel = pose_trans(rot_end, scoop_start_rel)

  	scoop_start_pose = pose_trans(p_center, scoop_start_rel)
  	scoop_via_pose = pose_trans(p_center, scoop_via_rel)
  	scoop_end_pose = pose_trans(p_center, scoop_end_rel)

  	movel(scoop_start_pose, a=0.5, v=0.3)
  	#movel(p_center, a=0.5, v=1.0)
  	#sleep(5.0)

  	if (level<90.0):
  		Rotate()
  	end

  	#movec(scoop_via_pose, scoop_end_pose, a=0.03, v=0.05)
  	movec(scoop_via_pose, scoop_end_pose, a=0.03, v=0.02)
  	#movel(pose_trans(get_actual_tcp_pose(), p[0,0,0,0,0,deg2rad(90.0)]), a=0.03, v=0.05)
  	sleep(1.0)
  	local ry_deg = map_tilt_to_ry_deg(angle_deg)
  	local ry = deg2rad(ry_deg)
  	local end_rel = pose_trans(pose_inv(p_center), scoop_end_pose)
  	local end_rel_tilted = pose_trans(end_rel, p[0, 0, 0, 0, ry, 0])
  	global tilted_pose_in_base = pose_trans(p_center, p[0,correction_y,correction_z,end_rel_tilted[3],end_rel_tilted[4], end_rel_tilted[5]])
  	global tilted_pose_in_base = pose_trans(tilted_pose_in_base, p[0, 0, spatula_len, 0, 0, 0])

  	if (Pow_name == "lactose_fine" or Pow_name == "Magnesium_sterate"):
  		tilt_send((angle_deg+5))
  	end
  	movel(tilted_pose_in_base, a=0.03, v=0.1)

  	if (Pow_name == "lactose_fine" or Pow_name == "Magnesium_sterate"):
  		tilt_send((angle_deg-5))
  	end

  	if (spatula=="spatula_flat_S" or spatula=="spatula_S"):
  		vibration_3()
  	else:
  		set_analog_out(0, vibration_voltage)
  	end
  	if (Pow_name=="Mannitol" or Pow_name =="NaCl"):
  		local n=1.4
  	else:
  		local n=1.5
  	end
  	local ry_level = deg2rad(ry_deg/n)
  	local end_rel_tilted_level = pose_trans(end_rel, p[0, 0, 0, 0, ry_level, 0])
  	local level_tilted_pose_in_base = pose_trans(p_center, p[0,correction_y,correction_z,end_rel_tilted_level[3],end_rel_tilted_level[4], end_rel_tilted_level[5]])
  	local level_tilted_pose_in_base = pose_trans(level_tilted_pose_in_base, p[0, 0, spatula_len, 0, 0, 0])

  	movel(level_tilted_pose_in_base, a=0.03, v=0.1)
  	#if (level>70.0):
  		#sleep(1.0)
  	#end
  	sleep(1.0)
  	#sleep(vibration_time)

  	movel(tilted_pose_in_base, a=0.03, v=0.1)
  	set_analog_out(0, 0.0)

  	tilt_pose_rel = pose_trans(pose_inv(p_center), tilted_pose_in_base)

  	lifted_pose_rel = pose_trans(lift_offset, tilt_pose_rel)

  	global lifted_pose = pose_trans(p_center, lifted_pose_rel)
  	movel(lifted_pose, a=0.03, v=0.1)
  	CCW_Rotate()
  end


  def center_pose():
  	trans_rel = p[-0.005, 0.05, -0.015, 0, 0, 0]

  	p_translated = pose_trans(place_pose, trans_rel)
  	cx = p_translated[0]
  	cy = p_translated[1]
  	cz = p_translated[2]

  	global p_center_vertical = p[cx,cy,cz, 0, 0, 4.09]

  	#movej(p_center_vertical, a =0.3, v =0.3)
  	return p_center_vertical
  end

  def updated_center_pose(p_center_vertical, angle_deg):
  	hinge_pose = pose_trans(p_center_vertical, p[0,0,-0.2,0,0,0])
  	local_rel = pose_trans(pose_inv(hinge_pose), p_center_vertical)

  	rot_tilt = p[0,0,0, -deg2rad(angle_deg),0,0]
  	local_rel_tilted = pose_trans(rot_tilt, local_rel)

  	global p_center = pose_trans(hinge_pose, local_rel_tilted)
  	return p_center
  end

  def tilt_send(angle):
  	socket_open("192.168.12.101", 80)
  	angle = 92.0 - angle
  	socket_send_string("Tilt,"+to_str(angle)+",0")
  	sync()
  	sleep(0.5)
  	socket_close()
  end

  def Motors_off():
  	socket_open("192.168.12.101", 80)
  	socket_send_string("Off,0,0")
  	sync()
  	sleep(0.5)
  	socket_close()
  end

  def Rotate():
  	socket_open("192.168.12.101", 80)
  	socket_send_string("FullRotation, 1, 2000")
  	sync()
  	sleep(0.5)
  	socket_close()
  end


  def CCW_Rotate():
  	socket_open("192.168.12.101", 80)
  	socket_send_string("FullRotation, -1, 2000")
  	sync()
  	sleep(0.5)
  	socket_close()
  end
  def tilt_to_home():
  	socket_open("192.168.12.101", 80)
  	socket_send_string("Home,0,0")
  	sync()
  	sleep(0.5)
  	socket_close()
  end



  $ 24 "Script: Weight_scale_socket.script"
  def get_weight():
  	socket_open("192.168.12.103", 3002)
  	sleep(0.2)
  	textmsg("socket opened successfully!")
  	socket_send_string("GET_WEIGHT")
  	sync()
  	sleep(0.5)
  	receiveFromServ = socket_read_ascii_float(6)
  	while (receiveFromServ[0] <1):
  		sleep(0.5)
  		receiveFromServ = socket_read_ascii_float(1)
  		textmsg("retrying read:", receiveFromServ)
  	end
  	textmsg("Received weight:", receiveFromServ[1])
  	socket_close()
  	sleep(0.2)
  	return receiveFromServ[1]
  end

  def tare_scale():
  	socket_open("192.168.12.103", 3002)
  	socket_send_string("TARE")
  	sleep(0.5)
  	socket_close()
  end

  def zero_scale():
  	socket_open("192.168.12.103", 3002)
  	socket_send_string("ZERO")
  	sleep(0.5)
  	socket_close()
  end

  def log_weight():
  	socket_open("192.168.12.103", 3002)
  	socket_send_string("LOG_WEIGHT")
  	sleep(0.5)
  	socket_close()
  end

  def send_target_info():
  	socket_open("192.168.12.103", 3002)
  	socket_send_string("SET_TARGET:" + to_str(target_weight))
  	sleep(0.2)
  	socket_close()
  end
  def send_powder_info():
  	socket_open("192.168.12.103", 3002)
  	socket_send_string("SET_POWDER:" + Pow_name)
  	sleep(0.2)
  	socket_close()
  end
  def send_spatula_info():
  	socket_open("192.168.12.103", 3002)
  	socket_send_string("SET_SPATULA:" + spatula)
  	sleep(0.2)
  	socket_close()
  end

  def send_level_info():
  	socket_open("192.168.12.103", 3002)
  	socket_send_string("SET_LEVEL:" + to_str(level))
  	sleep(0.2)
  	socket_close()
  end


  $ 25 "BeforeStarts"
  $ 26 "uLM"
  $ 27 "CMD_Stop≔ False "
  global CMD_Stop=  False
  $ 28 "CMD_Abort≔ False "
  global CMD_Abort=  False
  $ 29 "CMD_Clear≔ False "
  global CMD_Clear=  False
  $ 30 "STATE≔1"
  global STATE=1
  $ 31 "STATE_Info≔''"
  global STATE_Info=""
  $ 32 "ARM_Referenced≔ False "
  global ARM_Referenced=  False
  $ 33 "zero_ftsensor()"
  zero_ftsensor()
  $ 34 "poses init"
  $ 35 "PSE_A≔p[0,0,0,0,0,0]"
  global PSE_A=p[0,0,0,0,0,0]
  $ 36 "PSE_A_H≔p[0,0,0,0,0,0]"
  global PSE_A_H=p[0,0,0,0,0,0]
  $ 37 "PSE_R≔p[0,0,0,0,0,0]"
  global PSE_R=p[0,0,0,0,0,0]
  $ 38 "PSE_R_H≔p[0,0,0,0,0,0]"
  global PSE_R_H=p[0,0,0,0,0,0]
  $ 39 "PSE_T≔p[0,0,0,0,0,0]"
  global PSE_T=p[0,0,0,0,0,0]
  $ 40 "PSE_T_H≔p[0,0,0,0,0,0]"
  global PSE_T_H=p[0,0,0,0,0,0]
  $ 41 "PSE_C_E≔p[0,0,0,0,0,0]"
  global PSE_C_E=p[0,0,0,0,0,0]
  $ 42 "PSE_C_H≔p[0,0,0,0,0,0]"
  global PSE_C_H=p[0,0,0,0,0,0]
  $ 43 "PSE_C_S≔p[0,0,0,0,0,0]"
  global PSE_C_S=p[0,0,0,0,0,0]
  $ 44 "init_home_by_cartesian_pose(p[0,-0.400,0.300,0,0,0])"
  init_home_by_cartesian_pose(p[0,-0.400,0.300,0,0,0])
  $ 45 "Clearing"
  $ 46 "reset_error()"
  reset_error()
  $ 47 "reset_warning()"
  reset_warning()
  $ 48 "uGo"
  $ 50 "ugo_init( True ,'http://192.168.12.120:10001')"
  ugo_init(  True  ,"http://192.168.12.120:10001")
  $ 51 "ugo_update_outputs()"
  ugo_update_outputs()
  $ 52 "App"
  $ 53 "'ADD APPLICATION SPECIFIC COMMANDS'"
  # 'ADD APPLICATION SPECIFIC COMMANDS'
  $ 54 "Tools"
  $ 55 "OBJ_Picked≔gripper_has_object()"
  global OBJ_Picked=gripper_has_object()
  $ 56 "If OBJ_Picked"
  if (OBJ_Picked):
    # begin: URCap Program Node
    #   Source: Robotiq_Grippers, 3.17.0.105337, Robotiq Inc.
    #   Type: Gripper Activate
    $ 57 "Gripper Activate"

    kill rq_gripper_communication_thread
    rq_gripper_communication_thread_started = False
    rq_close_gripper_socket("1")
    rq_close_gripper_socket("2")
    rq_close_gripper_socket("3")
    rq_close_gripper_socket("4")

    rq_init_comm_if_connected(9, "1")
    rq_init_comm_if_connected(2, "2")
    rq_init_comm_if_connected(3, "3")
    rq_init_comm_if_connected(4, "4")
    rq_print_connected_grippers()
    rq_gripper_communication_thread = run rq_gripper_communication()

    while(not rq_gripper_communication_thread_started):
        sleep(0.008)
    end

    rq_set_max_current_for_all_grippers()

    reset_and_activate = False

    rq_activate_all_grippers(False)
    # end: URCap Program Node
  else:
    $ 58 "Else" "noBreak"
    # begin: URCap Program Node
    #   Source: Robotiq_Grippers, 3.17.0.105337, Robotiq Inc.
    #   Type: Gripper Activate
    $ 59 "Gripper Reset and Activate"

    kill rq_gripper_communication_thread
    rq_gripper_communication_thread_started = False
    rq_close_gripper_socket("1")
    rq_close_gripper_socket("2")
    rq_close_gripper_socket("3")
    rq_close_gripper_socket("4")

    rq_init_comm_if_connected(9, "1")
    rq_init_comm_if_connected(2, "2")
    rq_init_comm_if_connected(3, "3")
    rq_init_comm_if_connected(4, "4")
    rq_print_connected_grippers()
    rq_gripper_communication_thread = run rq_gripper_communication()

    while(not rq_gripper_communication_thread_started):
        sleep(0.008)
    end

    rq_set_max_current_for_all_grippers()

    reset_and_activate = True

